Fanuc KAREL source: kc00043.KL

-- PROVISIONAL review KL for V940-1; original PC SHA256 854ef012694a02a774c35aef2bd741709433435e694cfee8c48bb1002bd0c0fc
-- Incomplete behavior may be omitted. Consult companion uncertainty JSON. Do not deploy.
PROGRAM KC00043
%NOLOCKGROUP
BEGIN
  -- V9_ZERO_TABLE_METADATA_HINT layout=0002_ascii; no indexed target words; source/name/runtime held
  -- UNRESOLVED_PC offsets 5-35; opcodes 27,22,22,27,9D,31,7E,4A
  -- UNRESOLVED_PC offsets 40-44; opcodes 7F
END KC00043
